FUNCTION_BLOCK OUTPUT_HISTORY (* Offline identification prototype; see docs/adaptive/4diac-design.md *)
  (* Standard: 61499-2 *)
  (* Version 0.1, 2026-09-26, Guilherme *)
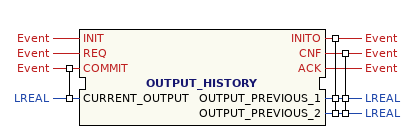
  EVENT_INPUT
    INIT;
    REQ;
    COMMIT WITH CURRENT_OUTPUT;
  END_EVENT
  EVENT_OUTPUT
    INITO WITH OUTPUT_PREVIOUS_1, OUTPUT_PREVIOUS_2;
    CNF WITH OUTPUT_PREVIOUS_1, OUTPUT_PREVIOUS_2;
    ACK;
  END_EVENT
  VAR_INPUT
    CURRENT_OUTPUT : LREAL;
  END_VAR
  VAR_OUTPUT
    OUTPUT_PREVIOUS_1 : LREAL;
    OUTPUT_PREVIOUS_2 : LREAL;
  END_VAR
  VAR
    H1 : LREAL;
    H2 : LREAL;
  END_VAR
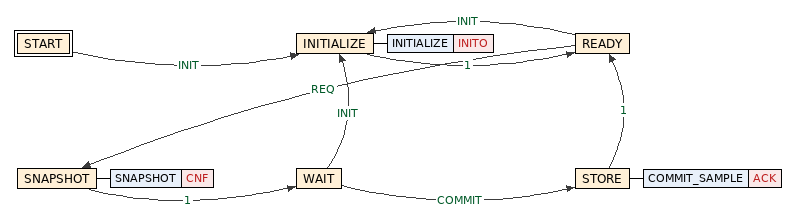
  EC_STATES
    START;
    INITIALIZE : INITIALIZE -> INITO;
    READY;
    SNAPSHOT : SNAPSHOT -> CNF;
    WAIT;
    STORE : COMMIT_SAMPLE -> ACK;
  END_STATES
  EC_TRANSITIONS
    START TO INITIALIZE := INIT;
    INITIALIZE TO READY := 1;
    READY TO INITIALIZE := INIT;
    READY TO SNAPSHOT := REQ;
    SNAPSHOT TO WAIT := 1;
    WAIT TO INITIALIZE := INIT;
    WAIT TO STORE := COMMIT;
    STORE TO READY := 1;
  END_TRANSITIONS
  ALGORITHM INITIALIZE IN ST:
H1 := 0.0;
H2 := 0.0;
OUTPUT_PREVIOUS_1 := 0.0;
OUTPUT_PREVIOUS_2 := 0.0;
  END_ALGORITHM
  ALGORITHM SNAPSHOT IN ST:
OUTPUT_PREVIOUS_1 := H1;
OUTPUT_PREVIOUS_2 := H2;
  END_ALGORITHM
  ALGORITHM COMMIT_SAMPLE IN ST:
H2 := H1;
H1 := CURRENT_OUTPUT;
  END_ALGORITHM
END_FUNCTION_BLOCK
